(* IEC 61131-3 sources: plc-st-coding-agent/progress/evidence/f14_v11_public_20261113/jobs/custom_deepseek-v4pro (part 4) *)

(* ---- public-medium-02.raw_candidate_01.st ---- *)
TYPE ST_AnalogChannel :
STRUCT
    enable : BOOL;
    hiLIM : REAL;
    loLIM : REAL;
    bipolar : BOOL;
    measuringMode : INT;
    retVal : WORD;
    outputValue : REAL;
END_STRUCT
END_TYPE

FUNCTION_BLOCK AnalogBatchProcessing
VAR_INPUT
    count : DINT;
END_VAR
VAR_INOUT
    analogValues : ARRAY[*] OF INT;
    channels : ARRAY[*] OF ST_AnalogChannel;
END_VAR
VAR
    tmp_i : DINT;
    tmp_process_count : DINT;
    tmp_analog_lower : DINT;
    tmp_channel_lower : DINT;
    tmp_analog_len : DINT;
    tmp_channel_len : DINT;
    tmp_raw : INT;
    tmp_raw_real : REAL;
    tmp_span : REAL;
    tmp_range : REAL;
END_VAR

(* ENGINEERING_CONTRACT
   Outputs:
   channels[].retVal : activation = enabled channel processed; retention = written only then; reset = none; priority = mode error before limit error; units: WORD.
   channels[].outputValue : activation = successful conversion only; retention = unchanged on skip/error/disabled; reset = none; units: REAL.
   Disabled channels: no writes.
   Mode 0 scaling boundaries: unipolar raw 0..27648 maps [loLIM,hiLIM], bipolar raw -27648..27648 maps [loLIM,hiLIM]; no clamping specified (PUB003).
   Mode 1/2 scale raw/10, raw/100 (PUB004, PUB005).
   Count represents ordinal positions from each array lower bound; caller valid 0..min lengths (PUB001). Cap invalid high count to available.
   Priority for invalid mode vs limit: invalid mode 16#8001 checked first, then limit 16#8002 (PUB006, PUB007).
*)

(* CONTRACT_RULES [] *)

tmp_analog_lower := LOWER_BOUND(analogValues, 1);
tmp_channel_lower := LOWER_BOUND(channels, 1);
tmp_analog_len := UPPER_BOUND(analogValues, 1) - tmp_analog_lower + 1;
tmp_channel_len := UPPER_BOUND(channels, 1) - tmp_channel_lower + 1;

IF count <= 0 THEN
    RETURN;
END_IF;

tmp_process_count := count;
IF tmp_process_count > tmp_analog_len THEN
    tmp_process_count := tmp_analog_len;
END_IF;
IF tmp_process_count > tmp_channel_len THEN
    tmp_process_count := tmp_channel_len;
END_IF;

FOR tmp_i := 0 TO tmp_process_count - 1 DO
    IF channels[tmp_channel_lower + tmp_i].enable THEN
        IF channels[tmp_channel_lower + tmp_i].measuringMode < 0 OR
           channels[tmp_channel_lower + tmp_i].measuringMode > 2 THEN
            channels[tmp_channel_lower + tmp_i].retVal := 16#8001;
        ELSIF channels[tmp_channel_lower + tmp_i].hiLIM <= channels[tmp_channel_lower + tmp_i].loLIM THEN
            channels[tmp_channel_lower + tmp_i].retVal := 16#8002;
        ELSE
            channels[tmp_channel_lower + tmp_i].retVal := 0;
            tmp_raw := analogValues[tmp_analog_lower + tmp_i];
            tmp_raw_real := TO_REAL(tmp_raw);
            CASE channels[tmp_channel_lower + tmp_i].measuringMode OF
                0:
                    tmp_span := channels[tmp_channel_lower + tmp_i].hiLIM - channels[tmp_channel_lower + tmp_i].loLIM;
                    IF channels[tmp_channel_lower + tmp_i].bipolar THEN
                        tmp_range := 55296.0;
                        channels[tmp_channel_lower + tmp_i].outputValue :=
                            channels[tmp_channel_lower + tmp_i].loLIM +
                            ((tmp_raw_real + 27648.0) / tmp_range) * tmp_span;
                    ELSE
                        tmp_range := 27648.0;
                        channels[tmp_channel_lower + tmp_i].outputValue :=
                            channels[tmp_channel_lower + tmp_i].loLIM +
                            (tmp_raw_real / tmp_range) * tmp_span;
                    END_IF
                1:
                    channels[tmp_channel_lower + tmp_i].outputValue := tmp_raw_real / 10.0;
                2:
                    channels[tmp_channel_lower + tmp_i].outputValue := tmp_raw_real / 100.0;
            END_CASE
        END_IF
    END_IF
END_FOR

END_FUNCTION_BLOCK

(* ---- public-medium-02.raw_candidate_02.st ---- *)
TYPE ST_AnalogChannel :
STRUCT
    enable : BOOL;
    hiLIM : REAL;
    loLIM : REAL;
    bipolar : BOOL;
    measuringMode : INT;
    retVal : WORD;
    outputValue : REAL;
END_STRUCT
END_TYPE;

FUNCTION_BLOCK AnalogBatchProcessing
VAR_INPUT
    count : DINT;
END_VAR
VAR_IN_OUT
    analogValues : ARRAY[*] OF INT;
    channels : ARRAY[*] OF ST_AnalogChannel;
END_VAR
VAR
    tmp_i : DINT;
    tmp_process_count : DINT;
    tmp_analog_lower : DINT;
    tmp_channel_lower : DINT;
    tmp_analog_len : DINT;
    tmp_channel_len : DINT;
    tmp_raw : INT;
    tmp_raw_real : REAL;
    tmp_span : REAL;
    tmp_range : REAL;
END_VAR

(* ENGINEERING_CONTRACT
   Outputs:
   channels[].retVal : activation = enabled channel processed; retention = written only then; reset = none; priority = mode error before limit error; units: WORD.
   channels[].outputValue : activation = successful conversion only; retention = unchanged on skip/error/disabled; reset = none; units: REAL.
   Disabled channels: no writes.
   Mode 0 scaling boundaries: unipolar raw 0..27648 maps [loLIM,hiLIM], bipolar raw -27648..27648 maps [loLIM,hiLIM]; no clamping specified (PUB003).
   Mode 1/2 scale raw/10, raw/100 (PUB004, PUB005).
   Count represents ordinal positions from each array lower bound; caller valid 0..min lengths (PUB001). Cap invalid high count to available.
   Priority for invalid mode vs limit: invalid mode 16#8001 checked first, then limit 16#8002 (PUB006, PUB007).
*)

(* CONTRACT_RULES [] *)

tmp_analog_lower := LOWER_BOUND(analogValues, 1);
tmp_channel_lower := LOWER_BOUND(channels, 1);
tmp_analog_len := UPPER_BOUND(analogValues, 1) - tmp_analog_lower + 1;
tmp_channel_len := UPPER_BOUND(channels, 1) - tmp_channel_lower + 1;

IF count <= 0 THEN
    RETURN;
END_IF;

tmp_process_count := count;
IF tmp_process_count > tmp_analog_len THEN
    tmp_process_count := tmp_analog_len;
END_IF;
IF tmp_process_count > tmp_channel_len THEN
    tmp_process_count := tmp_channel_len;
END_IF;

FOR tmp_i := 0 TO tmp_process_count - 1 DO
    IF channels[tmp_channel_lower + tmp_i].enable THEN
        IF channels[tmp_channel_lower + tmp_i].measuringMode < 0 OR
           channels[tmp_channel_lower + tmp_i].measuringMode > 2 THEN
            channels[tmp_channel_lower + tmp_i].retVal := 16#8001;
        ELSIF channels[tmp_channel_lower + tmp_i].hiLIM <= channels[tmp_channel_lower + tmp_i].loLIM THEN
            channels[tmp_channel_lower + tmp_i].retVal := 16#8002;
        ELSE
            channels[tmp_channel_lower + tmp_i].retVal := 0;
            tmp_raw := analogValues[tmp_analog_lower + tmp_i];
            tmp_raw_real := TO_REAL(tmp_raw);
            CASE channels[tmp_channel_lower + tmp_i].measuringMode OF
                0:
                    tmp_span := channels[tmp_channel_lower + tmp_i].hiLIM - channels[tmp_channel_lower + tmp_i].loLIM;
                    IF channels[tmp_channel_lower + tmp_i].bipolar THEN
                        tmp_range := 55296.0;
                        channels[tmp_channel_lower + tmp_i].outputValue :=
                            channels[tmp_channel_lower + tmp_i].loLIM +
                            ((tmp_raw_real + 27648.0) / tmp_range) * tmp_span;
                    ELSE
                        tmp_range := 27648.0;
                        channels[tmp_channel_lower + tmp_i].outputValue :=
                            channels[tmp_channel_lower + tmp_i].loLIM +
                            (tmp_raw_real / tmp_range) * tmp_span;
                    END_IF;
                1:
                    channels[tmp_channel_lower + tmp_i].outputValue := tmp_raw_real / 10.0;
                2:
                    channels[tmp_channel_lower + tmp_i].outputValue := tmp_raw_real / 100.0;
            END_CASE;
        END_IF;
    END_IF;
END_FOR;

END_FUNCTION_BLOCK

(* ---- public-medium-03.candidate_01.st ---- *)
FUNCTION_BLOCK FB
VAR_INPUT
    cyclicExecution : BOOL;
    trigger : BOOL;
    value : LREAL;
    windowSize : INT;
    reset : BOOL;
END_VAR
VAR_OUTPUT
    average : LREAL;
    windowSizeReached : BOOL;
    error : BOOL;
    status : WORD;
END_VAR
VAR
    trig_rt : R_TRIG;
    buf : ARRAY[0..99] OF LREAL;
    head : INT := 0;
    count : INT := 0;
    n : INT;
    i : INT;
    idx : INT;
    do_update : BOOL;
    tmp_sum : LREAL;
    tmp_window_valid : BOOL;
END_VAR

(* ENGINEERING_CONTRACT
   - average: LREAL, updated only on new value read (cyclic scan or trigger rising edge while cyclicExecution FALSE);
     reset clears to 0.0. Unit: input value unit.
   - windowSizeReached: BOOL, TRUE iff count >= windowSize and window valid; reset clears; invalid window sets FALSE.
   - error/status: combinational; invalid window (windowSize < 1 or > 100) sets error TRUE, status 16#8200;
     otherwise error FALSE, status 16#0000.
   - reset has priority over read; invalid window blocks read and overrides status; no latch.
   - trigger rising edges are ignored while cyclicExecution TRUE.
   - circular buffer capacity 100; changing windowSize does not clear buffer.
*)
(* CONTRACT_RULES [] *)

trig_rt(CLK := trigger);
tmp_window_valid := (windowSize >= 1) AND (windowSize <= 100);

IF reset THEN
    head := 0;
    count := 0;
    average := 0.0;
    windowSizeReached := FALSE;

    IF tmp_window_valid THEN
        error := FALSE;
        status := WORD#16#0000;
    ELSE
        error := TRUE;
        status := WORD#16#8200;
    END_IF;
    RETURN;

ELSIF NOT tmp_window_valid THEN
    error := TRUE;
    status := WORD#16#8200;
    average := 0.0;
    windowSizeReached := FALSE;
    RETURN;

ELSE
    error := FALSE;
    status := WORD#16#0000;
    windowSizeReached := (count >= windowSize);

    do_update := FALSE;
    IF cyclicExecution THEN
        do_update := TRUE;
    ELSIF trig_rt.Q THEN
        do_update := TRUE;
    END_IF;

    IF do_update THEN
        buf[head] := value;
        head := (head + 1) MOD 100;
        IF count < 100 THEN
            count := count + 1;
        END_IF;

        n := count;
        IF n > windowSize THEN
            n := windowSize;
        END_IF;

        IF n = 0 THEN
            average := 0.0;
        ELSE
            tmp_sum := 0.0;
            FOR i := 0 TO n - 1 DO
                idx := (head - n + i) MOD 100;
                IF idx < 0 THEN
                    idx := idx + 100;
                END_IF;
                tmp_sum := tmp_sum + buf[idx];
            END_FOR;
            average := tmp_sum / INT_TO_LREAL(n);
        END_IF;

        windowSizeReached := (count >= windowSize);
    END_IF;
END_IF;

END_FUNCTION_BLOCK

(* ---- public-medium-03.raw_candidate_01.st ---- *)
FUNCTION_BLOCK FB
VAR_INPUT
    cyclicExecution : BOOL;
    trigger : BOOL;
    value : LREAL;
    windowSize : INT;
    reset : BOOL;
END_VAR
VAR_OUTPUT
    average : LREAL;
    windowSizeReached : BOOL;
    error : BOOL;
    status : WORD;
END_VAR
VAR
    trig_rt : R_TRIG;
    buf : ARRAY[0..99] OF LREAL;
    head : INT := 0;
    count : INT := 0;
    n : INT;
    i : INT;
    idx : INT;
    do_update : BOOL;
    tmp_sum : LREAL;
    tmp_window_valid : BOOL;
END_VAR

(* ENGINEERING_CONTRACT
   - average: LREAL, updated only on new value read (cyclic scan or trigger rising edge while cyclicExecution FALSE);
     reset clears to 0.0. Unit: input value unit.
   - windowSizeReached: BOOL, TRUE iff count >= windowSize and window valid; reset clears; invalid window sets FALSE.
   - error/status: combinational; invalid window (windowSize < 1 or > 100) sets error TRUE, status 16#8200;
     otherwise error FALSE, status 16#0000.
   - reset has priority over read; invalid window blocks read and overrides status; no latch.
   - trigger rising edges are ignored while cyclicExecution TRUE.
   - circular buffer capacity 100; changing windowSize does not clear buffer.
*)
(* CONTRACT_RULES [] *)

trig_rt(CLK := trigger);
tmp_window_valid := (windowSize >= 1) AND (windowSize <= 100);

IF reset THEN
    head := 0;
    count := 0;
    average := 0.0;
    windowSizeReached := FALSE;

    IF tmp_window_valid THEN
        error := FALSE;
        status := WORD#16#0000;
    ELSE
        error := TRUE;
        status := WORD#16#8200;
    END_IF;
    RETURN;

ELSIF NOT tmp_window_valid THEN
    error := TRUE;
    status := WORD#16#8200;
    average := 0.0;
    windowSizeReached := FALSE;
    RETURN;

ELSE
    error := FALSE;
    status := WORD#16#0000;
    windowSizeReached := (count >= windowSize);

    do_update := FALSE;
    IF cyclicExecution THEN
        do_update := TRUE;
    ELSIF trig_rt.Q THEN
        do_update := TRUE;
    END_IF;

    IF do_update THEN
        buf[head] := value;
        head := (head + 1) MOD 100;
        IF count < 100 THEN
            count := count + 1;
        END_IF;

        n := count;
        IF n > windowSize THEN
            n := windowSize;
        END_IF;

        IF n = 0 THEN
            average := 0.0;
        ELSE
            tmp_sum := 0.0;
            FOR i := 0 TO n - 1 DO
                idx := (head - n + i) MOD 100;
                IF idx < 0 THEN
                    idx := idx + 100;
                END_IF;
                tmp_sum := tmp_sum + buf[idx];
            END_FOR;
            average := tmp_sum / INT_TO_LREAL(n);
        END_IF;

        windowSizeReached := (count >= windowSize);
    END_IF;
END_IF;

END_FUNCTION_BLOCK

(* ---- public-medium-04.candidate_01.st ---- *)
FUNCTION_BLOCK FB_TemperatureControl
VAR_INPUT
    TemperatureSensorInput : REAL;
    SetTemperature : REAL;
END_VAR
VAR_OUTPUT
    CurrentTemperature : REAL;
    SetTempDisplay : REAL;
    HeaterStatus : BOOL;
    OverheatProtection : BOOL;
    HeaterOutput : BOOL;
END_VAR
VAR
    tmp_sensor_fault : BOOL;
    tmp_heat_allowed : BOOL;
    tmp_overheat_active : BOOL;
    tmp_heat_on_timer : TON;
    tmp_cooldown_timer : TON;
    tmp_heat_limit : TIME := T#5001MS;  (* strictly > 5 s continuous heating *)
    tmp_cooldown_limit : TIME := T#3S;
END_VAR

(*
ENGINEERING_CONTRACT
- CurrentTemperature/SetTempDisplay: combinational echoes, raw units.
- HeaterOutput: on when sensor valid, no overheat, sensor < set;
  off when sensor >= set, sensor fault, or overheat. Equal is off.
- OverheatProtection: latched TRUE on continuous heater on >5s; auto clear after 3s cooldown.
- HeaterStatus: echo of HeaterOutput.
- Sensor fault: <0.0 or >100.0. Fault and overheat force heater off.
- Unspecified: equal setpoint and reset after cooldown interpreted as above.
- PUB001-PUB008.
*)

(* CONTRACT_RULES [] *)

tmp_sensor_fault := (TemperatureSensorInput < 0.0) OR (TemperatureSensorInput > 100.0);

tmp_heat_allowed := (NOT tmp_sensor_fault)
                    AND (NOT tmp_overheat_active)
                    AND (TemperatureSensorInput < SetTemperature);

tmp_heat_on_timer(IN := tmp_heat_allowed, PT := tmp_heat_limit);

IF tmp_heat_on_timer.Q THEN
    tmp_overheat_active := TRUE;
END_IF;

tmp_cooldown_timer(IN := tmp_overheat_active, PT := tmp_cooldown_limit);

IF tmp_cooldown_timer.Q THEN
    tmp_overheat_active := FALSE;
END_IF;

HeaterOutput := (NOT tmp_sensor_fault)
                AND (NOT tmp_overheat_active)
                AND (TemperatureSensorInput < SetTemperature);

HeaterStatus := HeaterOutput;
OverheatProtection := tmp_overheat_active;
CurrentTemperature := TemperatureSensorInput;
SetTempDisplay := SetTemperature;

END_FUNCTION_BLOCK

(* ---- public-medium-04.candidate_02.st ---- *)
FUNCTION_BLOCK FB_TemperatureControl
VAR_INPUT
    TemperatureSensorInput : REAL;
    SetTemperature : REAL;
END_VAR
VAR_OUTPUT
    CurrentTemperature : REAL;
    SetTempDisplay : REAL;
    HeaterStatus : BOOL;
    OverheatProtection : BOOL;
    HeaterOutput : BOOL;
END_VAR
VAR
    tmp_sensor_fault : BOOL;
    tmp_heat_allowed : BOOL;
    tmp_overheat_active : BOOL;
    tmp_heat_on_timer : TON;
    tmp_cooldown_timer : TON;
    tmp_heat_limit : TIME := T#5001MS;  (* strictly > 5 s continuous heating *)
    tmp_cooldown_limit : TIME := T#3S;
END_VAR

(*
ENGINEERING_CONTRACT
- CurrentTemperature/SetTempDisplay: combinational echoes, raw units.
- HeaterOutput: on when sensor valid, no overheat, sensor < set;
  off when sensor >= set, sensor fault, or overheat. Equal is off.
- OverheatProtection: latched TRUE on continuous heater on >5s; auto clear after 3s cooldown.
- HeaterStatus: echo of HeaterOutput.
- Sensor fault: <0.0 or >100.0. Fault and overheat force heater off.
- Equal setpoint and reset after cooldown interpreted as above.
- Heat timer starts in same scan as heater is newly enabled; heat trip starts cooldown in same scan.
- PUB001-PUB008.
*)

(* CONTRACT_RULES [] *)

tmp_sensor_fault := (TemperatureSensorInput < 0.0) OR (TemperatureSensorInput > 100.0);

(* Process cooldown for any currently active overheat before computing heater command *)
tmp_cooldown_timer(IN := tmp_overheat_active, PT := tmp_cooldown_limit);
IF tmp_cooldown_timer.Q THEN
    tmp_overheat_active := FALSE;
END_IF;

tmp_heat_allowed := (NOT tmp_sensor_fault) AND (NOT tmp_overheat_active) AND (TemperatureSensorInput < SetTemperature);
HeaterOutput := tmp_heat_allowed;

tmp_heat_on_timer(IN := HeaterOutput, PT := tmp_heat_limit);
IF tmp_heat_on_timer.Q THEN
    tmp_overheat_active := TRUE;
    HeaterOutput := FALSE;
    (* Start cooldown timer on the same scan as the overheat trip *)
    tmp_cooldown_timer(IN := TRUE, PT := tmp_cooldown_limit);
END_IF;

HeaterStatus := HeaterOutput;
OverheatProtection := tmp_overheat_active;
CurrentTemperature := TemperatureSensorInput;
SetTempDisplay := SetTemperature;

END_FUNCTION_BLOCK

(* ---- public-medium-04.candidate_03.st ---- *)
FUNCTION_BLOCK FB_TemperatureControl
VAR_INPUT
    TemperatureSensorInput : REAL;
    SetTemperature : REAL;
END_VAR
VAR_OUTPUT
    CurrentTemperature : REAL;
    SetTempDisplay : REAL;
    HeaterStatus : BOOL;
    OverheatProtection : BOOL;
    HeaterOutput : BOOL;
END_VAR
VAR
    tmp_sensor_fault : BOOL;
    tmp_heat_allowed : BOOL;
    tmp_overheat_active : BOOL;
    tmp_heat_on_timer : TON;
    tmp_cooldown_timer : TON;
    tmp_heat_limit : TIME := T#5001MS;  (* strictly more than 5 s continuous heating *)
    tmp_cooldown_limit : TIME := T#3S;
END_VAR

(*
ENGINEERING_CONTRACT
- CurrentTemperature/SetTempDisplay are combinational echoes of the inputs.
- Sensor fault when input < 0.0 or > 100.0; fault forces heater off.
- HeaterOutput is on only when sensor valid, overheat protection inactive,
  and TemperatureSensorInput < SetTemperature. Equal setpoint is off.
- OverheatProtection latches when continuous heater-on time exceeds 5 s,
  and clears after a 3 s cooldown. Cooldown and same-scan reactivation are
  evaluated so clearing protection allows heater and its timer in the same scan.
- HeaterStatus follows HeaterOutput.
*)

(* CONTRACT_RULES [] *)

tmp_sensor_fault := (TemperatureSensorInput < 0.0) OR (TemperatureSensorInput > 100.0);

(* Evaluate cooldown first so a completed cooldown can lift protection
   and permit heater startup during this same invocation. *)
tmp_cooldown_timer(IN := tmp_overheat_active, PT := tmp_cooldown_limit);
IF tmp_cooldown_timer.Q THEN
    tmp_overheat_active := FALSE;
END_IF;

tmp_heat_allowed := (NOT tmp_sensor_fault)
                    AND (NOT tmp_overheat_active)
                    AND (TemperatureSensorInput < SetTemperature);

tmp_heat_on_timer(IN := tmp_heat_allowed, PT := tmp_heat_limit);

IF tmp_heat_on_timer.Q THEN
    tmp_overheat_active := TRUE;
    (* Start cooldown in the same scan when the overheat latch occurs. *)
    tmp_cooldown_timer(IN := TRUE, PT := tmp_cooldown_limit);
END_IF;

HeaterOutput := (NOT tmp_sensor_fault)
                AND (NOT tmp_overheat_active)
                AND (TemperatureSensorInput < SetTemperature);

HeaterStatus := HeaterOutput;
OverheatProtection := tmp_overheat_active;
CurrentTemperature := TemperatureSensorInput;
SetTempDisplay := SetTemperature;

END_FUNCTION_BLOCK

(* ---- public-medium-04.candidate_04.st ---- *)
FUNCTION_BLOCK FB_TemperatureControl
VAR_INPUT
    TemperatureSensorInput : REAL;
    SetTemperature : REAL;
END_VAR
VAR_OUTPUT
    CurrentTemperature : REAL;
    SetTempDisplay : REAL;
    HeaterStatus : BOOL;
    OverheatProtection : BOOL;
    HeaterOutput : BOOL;
END_VAR
VAR
    tmp_sensor_fault : BOOL;
    tmp_heat_allowed : BOOL;
    tmp_overheat_active : BOOL;
    tmp_heat_on_timer : TON;
    tmp_cooldown_timer : TON;
    tmp_heat_limit : TIME := T#5001MS;  (* strictly > 5 s continuous heating *)
    tmp_cooldown_limit : TIME := T#3S;
END_VAR

(*
ENGINEERING_CONTRACT
- CurrentTemperature/SetTempDisplay: combinational echoes, raw units.
- HeaterOutput: on when sensor valid, no overheat, sensor < set;
  off when sensor >= set, sensor fault, or overheat. Equal is off.
- OverheatProtection: latched TRUE on continuous heater on >5s; auto clear after 3s cooldown.
- HeaterStatus: echo of HeaterOutput.
- Sensor fault: <0.0 or >100.0. Fault and overheat force heater off.
- Unspecified: equal setpoint and reset after cooldown interpreted as above.
- PUB001-PUB008.
*)

(* CONTRACT_RULES [] *)

tmp_sensor_fault := (TemperatureSensorInput < 0.0) OR (TemperatureSensorInput > 100.0);

(* Cooldown logic first: if overheat is active and cooldown elapsed, clear it. *)
tmp_cooldown_timer(IN := tmp_overheat_active, PT := tmp_cooldown_limit);
IF tmp_cooldown_timer.Q THEN
    tmp_overheat_active := FALSE;
END_IF;

(* Recompute heater allowed using possibly updated overheat state. *)
tmp_heat_allowed := (NOT tmp_sensor_fault)
                    AND (NOT tmp_overheat_active)
                    AND (TemperatureSensorInput < SetTemperature);

(* Run heat timer after cooldown so it starts immediately when heater becomes allowed. *)
tmp_heat_on_timer(IN := tmp_heat_allowed, PT := tmp_heat_limit);
IF tmp_heat_on_timer.Q THEN
    tmp_overheat_active := TRUE;
END_IF;

HeaterOutput := (NOT tmp_sensor_fault)
                AND (NOT tmp_overheat_active)
                AND (TemperatureSensorInput < SetTemperature);

HeaterStatus := HeaterOutput;
OverheatProtection := tmp_overheat_active;
CurrentTemperature := TemperatureSensorInput;
SetTempDisplay := SetTemperature;

END_FUNCTION_BLOCK

(* ---- public-medium-04.raw_candidate_01.st ---- *)
FUNCTION_BLOCK FB_TemperatureControl
VAR_INPUT
    TemperatureSensorInput : REAL;
    SetTemperature : REAL;
END_VAR
VAR_OUTPUT
    CurrentTemperature : REAL;
    SetTempDisplay : REAL;
    HeaterStatus : BOOL;
    OverheatProtection : BOOL;
    HeaterOutput : BOOL;
END_VAR
VAR
    tmp_sensor_fault : BOOL;
    tmp_heat_allowed : BOOL;
    tmp_overheat_active : BOOL;
    tmp_heat_on_timer : TON;
    tmp_cooldown_timer : TON;
    tmp_heat_limit : TIME := T#5001MS;  (* strictly > 5 s continuous heating *)
    tmp_cooldown_limit : TIME := T#3S;
END_VAR

(*
ENGINEERING_CONTRACT
- CurrentTemperature/SetTempDisplay: combinational echoes, raw units.
- HeaterOutput: on when sensor valid, no overheat, sensor < set;
  off when sensor >= set, sensor fault, or overheat. Equal is off.
- OverheatProtection: latched TRUE on continuous heater on >5s; auto clear after 3s cooldown.
- HeaterStatus: echo of HeaterOutput.
- Sensor fault: <0.0 or >100.0. Fault and overheat force heater off.
- Unspecified: equal setpoint and reset after cooldown interpreted as above.
- PUB001-PUB008.
*)

(* CONTRACT_RULES [] *)

tmp_sensor_fault := (TemperatureSensorInput < 0.0) OR (TemperatureSensorInput > 100.0);

tmp_heat_allowed := (NOT tmp_sensor_fault)
                    AND (NOT tmp_overheat_active)
                    AND (TemperatureSensorInput < SetTemperature);

tmp_heat_on_timer(IN := tmp_heat_allowed, PT := tmp_heat_limit);

IF tmp_heat_on_timer.Q THEN
    tmp_overheat_active := TRUE;
END_IF;

tmp_cooldown_timer(IN := tmp_overheat_active, PT := tmp_cooldown_limit);

IF tmp_cooldown_timer.Q THEN
    tmp_overheat_active := FALSE;
END_IF;

HeaterOutput := (NOT tmp_sensor_fault)
                AND (NOT tmp_overheat_active)
                AND (TemperatureSensorInput < SetTemperature);

HeaterStatus := HeaterOutput;
OverheatProtection := tmp_overheat_active;
CurrentTemperature := TemperatureSensorInput;
SetTempDisplay := SetTemperature;

END_FUNCTION_BLOCK

(* ---- public-medium-04.raw_candidate_02.st ---- *)
FUNCTION_BLOCK FB_TemperatureControl
VAR_INPUT
    TemperatureSensorInput : REAL;
    SetTemperature : REAL;
END_VAR
VAR_OUTPUT
    CurrentTemperature : REAL;
    SetTempDisplay : REAL;
    HeaterStatus : BOOL;
    OverheatProtection : BOOL;
    HeaterOutput : BOOL;
END_VAR
VAR
    tmp_sensor_fault : BOOL;
    tmp_heat_allowed : BOOL;
    tmp_overheat_active : BOOL;
    tmp_heat_on_timer : TON;
    tmp_cooldown_timer : TON;
    tmp_heat_limit : TIME := T#5001MS;  (* strictly > 5 s continuous heating *)
    tmp_cooldown_limit : TIME := T#3S;
END_VAR

(*
ENGINEERING_CONTRACT
- CurrentTemperature/SetTempDisplay: combinational echoes, raw units.
- HeaterOutput: on when sensor valid, no overheat, sensor < set;
  off when sensor >= set, sensor fault, or overheat. Equal is off.
- OverheatProtection: latched TRUE on continuous heater on >5s; auto clear after 3s cooldown.
- HeaterStatus: echo of HeaterOutput.
- Sensor fault: <0.0 or >100.0. Fault and overheat force heater off.
- Equal setpoint and reset after cooldown interpreted as above.
- Heat timer starts in same scan as heater is newly enabled; heat trip starts cooldown in same scan.
- PUB001-PUB008.
*)

(* CONTRACT_RULES [] *)

tmp_sensor_fault := (TemperatureSensorInput < 0.0) OR (TemperatureSensorInput > 100.0);

(* Process cooldown for any currently active overheat before computing heater command *)
tmp_cooldown_timer(IN := tmp_overheat_active, PT := tmp_cooldown_limit);
IF tmp_cooldown_timer.Q THEN
    tmp_overheat_active := FALSE;
END_IF;

tmp_heat_allowed := (NOT tmp_sensor_fault) AND (NOT tmp_overheat_active) AND (TemperatureSensorInput < SetTemperature);
HeaterOutput := tmp_heat_allowed;

tmp_heat_on_timer(IN := HeaterOutput, PT := tmp_heat_limit);
IF tmp_heat_on_timer.Q THEN
    tmp_overheat_active := TRUE;
    HeaterOutput := FALSE;
    (* Start cooldown timer on the same scan as the overheat trip *)
    tmp_cooldown_timer(IN := TRUE, PT := tmp_cooldown_limit);
END_IF;

HeaterStatus := HeaterOutput;
OverheatProtection := tmp_overheat_active;
CurrentTemperature := TemperatureSensorInput;
SetTempDisplay := SetTemperature;

END_FUNCTION_BLOCK

(* ---- public-medium-04.raw_candidate_03.st ---- *)
FUNCTION_BLOCK FB_TemperatureControl
VAR_INPUT
    TemperatureSensorInput : REAL;
    SetTemperature : REAL;
END_VAR
VAR_OUTPUT
    CurrentTemperature : REAL;
    SetTempDisplay : REAL;
    HeaterStatus : BOOL;
    OverheatProtection : BOOL;
    HeaterOutput : BOOL;
END_VAR
VAR
    tmp_sensor_fault : BOOL;
    tmp_heat_allowed : BOOL;
    tmp_overheat_active : BOOL;
    tmp_heat_on_timer : TON;
    tmp_cooldown_timer : TON;
    tmp_heat_limit : TIME := T#5001MS;  (* strictly more than 5 s continuous heating *)
    tmp_cooldown_limit : TIME := T#3S;
END_VAR

(*
ENGINEERING_CONTRACT
- CurrentTemperature/SetTempDisplay are combinational echoes of the inputs.
- Sensor fault when input < 0.0 or > 100.0; fault forces heater off.
- HeaterOutput is on only when sensor valid, overheat protection inactive,
  and TemperatureSensorInput < SetTemperature. Equal setpoint is off.
- OverheatProtection latches when continuous heater-on time exceeds 5 s,
  and clears after a 3 s cooldown. Cooldown and same-scan reactivation are
  evaluated so clearing protection allows heater and its timer in the same scan.
- HeaterStatus follows HeaterOutput.
*)

(* CONTRACT_RULES [] *)

tmp_sensor_fault := (TemperatureSensorInput < 0.0) OR (TemperatureSensorInput > 100.0);

(* Evaluate cooldown first so a completed cooldown can lift protection
   and permit heater startup during this same invocation. *)
tmp_cooldown_timer(IN := tmp_overheat_active, PT := tmp_cooldown_limit);
IF tmp_cooldown_timer.Q THEN
    tmp_overheat_active := FALSE;
END_IF;

tmp_heat_allowed := (NOT tmp_sensor_fault)
                    AND (NOT tmp_overheat_active)
                    AND (TemperatureSensorInput < SetTemperature);

tmp_heat_on_timer(IN := tmp_heat_allowed, PT := tmp_heat_limit);

IF tmp_heat_on_timer.Q THEN
    tmp_overheat_active := TRUE;
    (* Start cooldown in the same scan when the overheat latch occurs. *)
    tmp_cooldown_timer(IN := TRUE, PT := tmp_cooldown_limit);
END_IF;

HeaterOutput := (NOT tmp_sensor_fault)
                AND (NOT tmp_overheat_active)
                AND (TemperatureSensorInput < SetTemperature);

HeaterStatus := HeaterOutput;
OverheatProtection := tmp_overheat_active;
CurrentTemperature := TemperatureSensorInput;
SetTempDisplay := SetTemperature;

END_FUNCTION_BLOCK

(* ---- public-medium-04.raw_candidate_04.st ---- *)
FUNCTION_BLOCK FB_TemperatureControl
VAR_INPUT
    TemperatureSensorInput : REAL;
    SetTemperature : REAL;
END_VAR
VAR_OUTPUT
    CurrentTemperature : REAL;
    SetTempDisplay : REAL;
    HeaterStatus : BOOL;
    OverheatProtection : BOOL;
    HeaterOutput : BOOL;
END_VAR
VAR
    tmp_sensor_fault : BOOL;
    tmp_heat_allowed : BOOL;
    tmp_overheat_active : BOOL;
    tmp_heat_on_timer : TON;
    tmp_cooldown_timer : TON;
    tmp_heat_limit : TIME := T#5001MS;  (* strictly > 5 s continuous heating *)
    tmp_cooldown_limit : TIME := T#3S;
END_VAR

(*
ENGINEERING_CONTRACT
- CurrentTemperature/SetTempDisplay: combinational echoes, raw units.
- HeaterOutput: on when sensor valid, no overheat, sensor < set;
  off when sensor >= set, sensor fault, or overheat. Equal is off.
- OverheatProtection: latched TRUE on continuous heater on >5s; auto clear after 3s cooldown.
- HeaterStatus: echo of HeaterOutput.
- Sensor fault: <0.0 or >100.0. Fault and overheat force heater off.
- Unspecified: equal setpoint and reset after cooldown interpreted as above.
- PUB001-PUB008.
*)

(* CONTRACT_RULES [] *)

tmp_sensor_fault := (TemperatureSensorInput < 0.0) OR (TemperatureSensorInput > 100.0);

(* Cooldown logic first: if overheat is active and cooldown elapsed, clear it. *)
tmp_cooldown_timer(IN := tmp_overheat_active, PT := tmp_cooldown_limit);
IF tmp_cooldown_timer.Q THEN
    tmp_overheat_active := FALSE;
END_IF;

(* Recompute heater allowed using possibly updated overheat state. *)
tmp_heat_allowed := (NOT tmp_sensor_fault)
                    AND (NOT tmp_overheat_active)
                    AND (TemperatureSensorInput < SetTemperature);

(* Run heat timer after cooldown so it starts immediately when heater becomes allowed. *)
tmp_heat_on_timer(IN := tmp_heat_allowed, PT := tmp_heat_limit);
IF tmp_heat_on_timer.Q THEN
    tmp_overheat_active := TRUE;
END_IF;

HeaterOutput := (NOT tmp_sensor_fault)
                AND (NOT tmp_overheat_active)
                AND (TemperatureSensorInput < SetTemperature);

HeaterStatus := HeaterOutput;
OverheatProtection := tmp_overheat_active;
CurrentTemperature := TemperatureSensorInput;
SetTempDisplay := SetTemperature;

END_FUNCTION_BLOCK

(* ---- public-medium-05.candidate_01.st ---- *)
(* ENGINEERING_CONTRACT
- Manual mode (Mode=FALSE): MotorForward set while ForwardButton AND NOT ReverseButton; MotorReverse set while ReverseButton AND NOT ForwardButton; simultaneous buttons deactivate both (PUB002).
- Automatic mode (Mode=TRUE): move_AB latch set by ButtonA R_TRIG while SensorA true; cleared when SensorB true. move_BC latch set by ButtonB R_TRIG while SensorB true; cleared when SensorC true.
- MotorForward = Mode AND (move_AB OR move_BC). MotorReverse is always FALSE in automatic mode (PUB003/PUB004).
- CompletionLight latch set by ButtonC R_TRIG while Mode=TRUE and SensorC true; held high; cleared when SensorC=FALSE regardless of Mode (PUB004).
- Same-scan priority: destination sensor clear wins over move set; simultaneous ForwardButton and ReverseButton -> both motor outputs FALSE.
*)

(* CONTRACT_RULES [] *)

FUNCTION_BLOCK ProductionLineControl
VAR_INPUT
    Mode : BOOL;
    ForwardButton : BOOL;
    ReverseButton : BOOL;
    SensorA : BOOL;
    SensorB : BOOL;
    SensorC : BOOL;
    ButtonA : BOOL;
    ButtonB : BOOL;
    ButtonC : BOOL;
END_VAR
VAR_OUTPUT
    MotorForward : BOOL;
    MotorReverse : BOOL;
    CompletionLight : BOOL;
END_VAR
VAR
    move_AB : BOOL := FALSE;
    move_BC : BOOL := FALSE;
    completion_latch : BOOL := FALSE;
    btnA_rt : R_TRIG;
    btnB_rt : R_TRIG;
    btnC_rt : R_TRIG;
END_VAR

btnA_rt(CLK := ButtonA);
btnB_rt(CLK := ButtonB);
btnC_rt(CLK := ButtonC);

IF Mode THEN
    IF btnA_rt.Q AND SensorA THEN
        move_AB := TRUE;
    END_IF;

    IF btnB_rt.Q AND SensorB THEN
        move_BC := TRUE;
    END_IF;

    IF btnC_rt.Q AND SensorC THEN
        completion_latch := TRUE;
    END_IF;
END_IF;

IF SensorB THEN
    move_AB := FALSE;
END_IF;

IF SensorC THEN
    move_BC := FALSE;
END_IF;

IF NOT SensorC THEN
    completion_latch := FALSE;
END_IF;

IF Mode THEN
    MotorForward := move_AB OR move_BC;
    MotorReverse := FALSE;
ELSE
    IF ForwardButton AND NOT ReverseButton THEN
        MotorForward := TRUE;
        MotorReverse := FALSE;
    ELSIF ReverseButton AND NOT ForwardButton THEN
        MotorForward := FALSE;
        MotorReverse := TRUE;
    ELSE
        MotorForward := FALSE;
        MotorReverse := FALSE;
    END_IF;
END_IF;

CompletionLight := completion_latch;

END_FUNCTION_BLOCK

(* ---- public-medium-05.candidate_02.st ---- *)
(* ENGINEERING_CONTRACT
- Manual mode (Mode=FALSE): MotorForward set while ForwardButton AND NOT ReverseButton; MotorReverse set while ReverseButton AND NOT ForwardButton; simultaneous buttons deactivate both (PUB002).
- Automatic mode (Mode=TRUE): move_AB latch set by ButtonA R_TRIG while SensorA true; cleared when SensorB true. move_BC latch set by ButtonB while SensorB true; cleared when SensorC true.
- MotorForward = Mode AND (move_AB OR move_BC). MotorReverse is always FALSE in automatic mode (PUB003/PUB004).
- CompletionLight latch set by ButtonC R_TRIG while Mode=TRUE and SensorC true; held high; cleared when SensorC=FALSE regardless of Mode (PUB004).
- Same-scan priority: destination sensor clear wins over move set; simultaneous ForwardButton and ReverseButton -> both motor outputs FALSE.
*)

(* CONTRACT_RULES [] *)

FUNCTION_BLOCK ProductionLineControl
VAR_INPUT
    Mode : BOOL;
    ForwardButton : BOOL;
    ReverseButton : BOOL;
    SensorA : BOOL;
    SensorB : BOOL;
    SensorC : BOOL;
    ButtonA : BOOL;
    ButtonB : BOOL;
    ButtonC : BOOL;
END_VAR
VAR_OUTPUT
    MotorForward : BOOL;
    MotorReverse : BOOL;
    CompletionLight : BOOL;
END_VAR
VAR
    move_AB : BOOL := FALSE;
    move_BC : BOOL := FALSE;
    completion_latch : BOOL := FALSE;
    btnA_rt : R_TRIG;
    btnB_rt : R_TRIG;
    btnC_rt : R_TRIG;
END_VAR

btnA_rt(CLK := ButtonA);
btnB_rt(CLK := ButtonB);
btnC_rt(CLK := ButtonC);

IF Mode THEN
    IF btnA_rt.Q AND SensorA THEN
        move_AB := TRUE;
    END_IF;

    IF ButtonB AND SensorB THEN
        move_BC := TRUE;
    END_IF;

    IF btnC_rt.Q AND SensorC THEN
        completion_latch := TRUE;
    END_IF;
END_IF;

IF SensorB THEN
    move_AB := FALSE;
END_IF;

IF SensorC THEN
    move_BC := FALSE;
END_IF;

IF NOT SensorC THEN
    completion_latch := FALSE;
END_IF;

IF Mode THEN
    MotorForward := move_AB OR move_BC;
    MotorReverse := FALSE;
ELSE
    IF ForwardButton AND NOT ReverseButton THEN
        MotorForward := TRUE;
        MotorReverse := FALSE;
    ELSIF ReverseButton AND NOT ForwardButton THEN
        MotorForward := FALSE;
        MotorReverse := TRUE;
    ELSE
        MotorForward := FALSE;
        MotorReverse := FALSE;
    END_IF;
END_IF;

CompletionLight := completion_latch;

END_FUNCTION_BLOCK

(* ---- public-medium-05.candidate_03.st ---- *)
(* ENGINEERING_CONTRACT
- Manual mode (Mode=FALSE): MotorForward set while ForwardButton AND NOT ReverseButton; MotorReverse set while ReverseButton AND NOT ForwardButton; simultaneous buttons deactivate both (PUB002).
- Automatic mode (Mode=TRUE): move_AB latch set by ButtonA R_TRIG while SensorA true; cleared when SensorB true. move_BC latch set by ButtonB while SensorB true; cleared when SensorC true.
- MotorForward = Mode AND (move_AB OR move_BC). MotorReverse is always FALSE in automatic mode (PUB003/PUB004).
- CompletionLight latch set by ButtonC R_TRIG while Mode=TRUE and SensorC true; held high; cleared when SensorC=FALSE regardless of Mode (PUB004).
- Same-scan priority: destination sensor clear wins over move set; simultaneous ForwardButton and ReverseButton -> both motor outputs FALSE.
*)

(* CONTRACT_RULES [] *)

FUNCTION_BLOCK ProductionLineControl
VAR_INPUT
    Mode : BOOL;
    ForwardButton : BOOL;
    ReverseButton : BOOL;
    SensorA : BOOL;
    SensorB : BOOL;
    SensorC : BOOL;
    ButtonA : BOOL;
    ButtonB : BOOL;
    ButtonC : BOOL;
END_VAR
VAR_OUTPUT
    MotorForward : BOOL;
    MotorReverse : BOOL;
    CompletionLight : BOOL;
END_VAR
VAR
    move_AB : BOOL := FALSE;
    move_BC : BOOL := FALSE;
    completion_latch : BOOL := FALSE;
    btnA_rt : R_TRIG;
    btnB_rt : R_TRIG;
    btnC_rt : R_TRIG;
END_VAR

btnA_rt(CLK := ButtonA);
btnB_rt(CLK := ButtonB);
btnC_rt(CLK := ButtonC);

IF Mode THEN
    IF btnA_rt.Q AND SensorA THEN
        move_AB := TRUE;
    END_IF;

    IF btnB_rt.Q AND SensorB THEN
        move_BC := TRUE;
    END_IF;

    IF btnC_rt.Q AND SensorC THEN
        completion_latch := TRUE;
    END_IF;
END_IF;

IF SensorB THEN
    move_AB := FALSE;
END_IF;

IF SensorC THEN
    move_BC := FALSE;
END_IF;

IF NOT SensorC THEN
    completion_latch := FALSE;
END_IF;

IF Mode THEN
    MotorForward := move_AB OR move_BC;
    MotorReverse := FALSE;
ELSE
    IF ForwardButton AND NOT ReverseButton THEN
        MotorForward := TRUE;
        MotorReverse := FALSE;
    ELSIF ReverseButton AND NOT ForwardButton THEN
        MotorForward := FALSE;
        MotorReverse := TRUE;
    ELSE
        MotorForward := FALSE;
        MotorReverse := FALSE;
    END_IF;
END_IF;

CompletionLight := completion_latch;

END_FUNCTION_BLOCK

(* ---- public-medium-05.candidate_04.st ---- *)
(* ENGINEERING_CONTRACT
- Manual mode (Mode=FALSE): MotorForward set while ForwardButton AND NOT ReverseButton; MotorReverse set while ReverseButton AND NOT ForwardButton; simultaneous buttons deactivate both (PUB002).
- Automatic mode (Mode=TRUE): move_AB latch set by ButtonA R_TRIG while SensorA true; cleared when SensorB true. move_BC latch set by ButtonB R_TRIG while SensorB true; cleared when SensorC true.
- MotorForward = Mode AND (move_AB OR move_BC). MotorReverse is always FALSE in automatic mode (PUB003/PUB004).
- CompletionLight latch set by ButtonC R_TRIG while Mode=TRUE and SensorC true; held high; cleared when SensorC=FALSE regardless of Mode (PUB004).
- Same-scan priority: destination sensor clear wins over move set; simultaneous ForwardButton and ReverseButton -> both motor outputs FALSE.
*)

(* CONTRACT_RULES [] *)

FUNCTION_BLOCK ProductionLineControl
VAR_INPUT
    Mode : BOOL;
    ForwardButton : BOOL;
    ReverseButton : BOOL;
    SensorA : BOOL;
    SensorB : BOOL;
    SensorC : BOOL;
    ButtonA : BOOL;
    ButtonB : BOOL;
    ButtonC : BOOL;
END_VAR
VAR_OUTPUT
    MotorForward : BOOL;
    MotorReverse : BOOL;
    CompletionLight : BOOL;
END_VAR
VAR
    move_AB : BOOL := FALSE;
    move_BC : BOOL := FALSE;
    completion_latch : BOOL := FALSE;
    btnA_rt : R_TRIG;
    btnB_rt : R_TRIG;
    btnC_rt : R_TRIG;
END_VAR

btnA_rt(CLK := ButtonA);
btnB_rt(CLK := ButtonB);
btnC_rt(CLK := ButtonC);

IF Mode THEN
    IF btnA_rt.Q AND SensorA THEN
        move_AB := TRUE;
    END_IF;

    IF btnB_rt.Q AND SensorB THEN
        move_BC := TRUE;
    END_IF;

    IF btnC_rt.Q AND SensorC THEN
        completion_latch := TRUE;
    END_IF;
END_IF;

IF SensorB THEN
    move_AB := FALSE;
END_IF;

IF SensorC THEN
    move_BC := FALSE;
END_IF;

IF NOT SensorC THEN
    completion_latch := FALSE;
END_IF;

IF Mode THEN
    MotorForward := move_AB OR move_BC;
    MotorReverse := FALSE;
ELSE
    IF ForwardButton AND NOT ReverseButton THEN
        MotorForward := TRUE;
        MotorReverse := FALSE;
    ELSIF ReverseButton AND NOT ForwardButton THEN
        MotorForward := FALSE;
        MotorReverse := TRUE;
    ELSE
        MotorForward := FALSE;
        MotorReverse := FALSE;
    END_IF;
END_IF;

CompletionLight := completion_latch;

END_FUNCTION_BLOCK

(* ---- public-medium-05.raw_candidate_01.st ---- *)
(* ENGINEERING_CONTRACT
- Manual mode (Mode=FALSE): MotorForward set while ForwardButton AND NOT ReverseButton; MotorReverse set while ReverseButton AND NOT ForwardButton; simultaneous buttons deactivate both (PUB002).
- Automatic mode (Mode=TRUE): move_AB latch set by ButtonA R_TRIG while SensorA true; cleared when SensorB true. move_BC latch set by ButtonB R_TRIG while SensorB true; cleared when SensorC true.
- MotorForward = Mode AND (move_AB OR move_BC). MotorReverse is always FALSE in automatic mode (PUB003/PUB004).
- CompletionLight latch set by ButtonC R_TRIG while Mode=TRUE and SensorC true; held high; cleared when SensorC=FALSE regardless of Mode (PUB004).
- Same-scan priority: destination sensor clear wins over move set; simultaneous ForwardButton and ReverseButton -> both motor outputs FALSE.
*)

(* CONTRACT_RULES [] *)

FUNCTION_BLOCK ProductionLineControl
VAR_INPUT
    Mode : BOOL;
    ForwardButton : BOOL;
    ReverseButton : BOOL;
    SensorA : BOOL;
    SensorB : BOOL;
    SensorC : BOOL;
    ButtonA : BOOL;
    ButtonB : BOOL;
    ButtonC : BOOL;
END_VAR
VAR_OUTPUT
    MotorForward : BOOL;
    MotorReverse : BOOL;
    CompletionLight : BOOL;
END_VAR
VAR
    move_AB : BOOL := FALSE;
    move_BC : BOOL := FALSE;
    completion_latch : BOOL := FALSE;
    btnA_rt : R_TRIG;
    btnB_rt : R_TRIG;
    btnC_rt : R_TRIG;
END_VAR

btnA_rt(CLK := ButtonA);
btnB_rt(CLK := ButtonB);
btnC_rt(CLK := ButtonC);

IF Mode THEN
    IF btnA_rt.Q AND SensorA THEN
        move_AB := TRUE;
    END_IF;

    IF btnB_rt.Q AND SensorB THEN
        move_BC := TRUE;
    END_IF;

    IF btnC_rt.Q AND SensorC THEN
        completion_latch := TRUE;
    END_IF;
END_IF;

IF SensorB THEN
    move_AB := FALSE;
END_IF;

IF SensorC THEN
    move_BC := FALSE;
END_IF;

IF NOT SensorC THEN
    completion_latch := FALSE;
END_IF;

IF Mode THEN
    MotorForward := move_AB OR move_BC;
    MotorReverse := FALSE;
ELSE
    IF ForwardButton AND NOT ReverseButton THEN
        MotorForward := TRUE;
        MotorReverse := FALSE;
    ELSIF ReverseButton AND NOT ForwardButton THEN
        MotorForward := FALSE;
        MotorReverse := TRUE;
    ELSE
        MotorForward := FALSE;
        MotorReverse := FALSE;
    END_IF;
END_IF;

CompletionLight := completion_latch;

END_FUNCTION_BLOCK

(* ---- public-medium-05.raw_candidate_02.st ---- *)
(* ENGINEERING_CONTRACT
- Manual mode (Mode=FALSE): MotorForward set while ForwardButton AND NOT ReverseButton; MotorReverse set while ReverseButton AND NOT ForwardButton; simultaneous buttons deactivate both (PUB002).
- Automatic mode (Mode=TRUE): move_AB latch set by ButtonA R_TRIG while SensorA true; cleared when SensorB true. move_BC latch set by ButtonB while SensorB true; cleared when SensorC true.
- MotorForward = Mode AND (move_AB OR move_BC). MotorReverse is always FALSE in automatic mode (PUB003/PUB004).
- CompletionLight latch set by ButtonC R_TRIG while Mode=TRUE and SensorC true; held high; cleared when SensorC=FALSE regardless of Mode (PUB004).
- Same-scan priority: destination sensor clear wins over move set; simultaneous ForwardButton and ReverseButton -> both motor outputs FALSE.
*)

(* CONTRACT_RULES [] *)

FUNCTION_BLOCK ProductionLineControl
VAR_INPUT
    Mode : BOOL;
    ForwardButton : BOOL;
    ReverseButton : BOOL;
    SensorA : BOOL;
    SensorB : BOOL;
    SensorC : BOOL;
    ButtonA : BOOL;
    ButtonB : BOOL;
    ButtonC : BOOL;
END_VAR
VAR_OUTPUT
    MotorForward : BOOL;
    MotorReverse : BOOL;
    CompletionLight : BOOL;
END_VAR
VAR
    move_AB : BOOL := FALSE;
    move_BC : BOOL := FALSE;
    completion_latch : BOOL := FALSE;
    btnA_rt : R_TRIG;
    btnB_rt : R_TRIG;
    btnC_rt : R_TRIG;
END_VAR

btnA_rt(CLK := ButtonA);
btnB_rt(CLK := ButtonB);
btnC_rt(CLK := ButtonC);

IF Mode THEN
    IF btnA_rt.Q AND SensorA THEN
        move_AB := TRUE;
    END_IF;

    IF ButtonB AND SensorB THEN
        move_BC := TRUE;
    END_IF;

    IF btnC_rt.Q AND SensorC THEN
        completion_latch := TRUE;
    END_IF;
END_IF;

IF SensorB THEN
    move_AB := FALSE;
END_IF;

IF SensorC THEN
    move_BC := FALSE;
END_IF;

IF NOT SensorC THEN
    completion_latch := FALSE;
END_IF;

IF Mode THEN
    MotorForward := move_AB OR move_BC;
    MotorReverse := FALSE;
ELSE
    IF ForwardButton AND NOT ReverseButton THEN
        MotorForward := TRUE;
        MotorReverse := FALSE;
    ELSIF ReverseButton AND NOT ForwardButton THEN
        MotorForward := FALSE;
        MotorReverse := TRUE;
    ELSE
        MotorForward := FALSE;
        MotorReverse := FALSE;
    END_IF;
END_IF;

CompletionLight := completion_latch;

END_FUNCTION_BLOCK

(* ---- public-medium-05.raw_candidate_03.st ---- *)
(* ENGINEERING_CONTRACT
- Manual mode (Mode=FALSE): MotorForward set while ForwardButton AND NOT ReverseButton; MotorReverse set while ReverseButton AND NOT ForwardButton; simultaneous buttons deactivate both (PUB002).
- Automatic mode (Mode=TRUE): move_AB latch set by ButtonA R_TRIG while SensorA true; cleared when SensorB true. move_BC latch set by ButtonB while SensorB true; cleared when SensorC true.
- MotorForward = Mode AND (move_AB OR move_BC). MotorReverse is always FALSE in automatic mode (PUB003/PUB004).
- CompletionLight latch set by ButtonC R_TRIG while Mode=TRUE and SensorC true; held high; cleared when SensorC=FALSE regardless of Mode (PUB004).
- Same-scan priority: destination sensor clear wins over move set; simultaneous ForwardButton and ReverseButton -> both motor outputs FALSE.
*)

(* CONTRACT_RULES [] *)

FUNCTION_BLOCK ProductionLineControl
VAR_INPUT
    Mode : BOOL;
    ForwardButton : BOOL;
    ReverseButton : BOOL;
    SensorA : BOOL;
    SensorB : BOOL;
    SensorC : BOOL;
    ButtonA : BOOL;
    ButtonB : BOOL;
    ButtonC : BOOL;
END_VAR
VAR_OUTPUT
    MotorForward : BOOL;
    MotorReverse : BOOL;
    CompletionLight : BOOL;
END_VAR
VAR
    move_AB : BOOL := FALSE;
    move_BC : BOOL := FALSE;
    completion_latch : BOOL := FALSE;
    btnA_rt : R_TRIG;
    btnB_rt : R_TRIG;
    btnC_rt : R_TRIG;
END_VAR

btnA_rt(CLK := ButtonA);
btnB_rt(CLK := ButtonB);
btnC_rt(CLK := ButtonC);

IF Mode THEN
    IF btnA_rt.Q AND SensorA THEN
        move_AB := TRUE;
    END_IF;

    IF btnB_rt.Q AND SensorB THEN
        move_BC := TRUE;
    END_IF;

    IF btnC_rt.Q AND SensorC THEN
        completion_latch := TRUE;
    END_IF;
END_IF;

IF SensorB THEN
    move_AB := FALSE;
END_IF;

IF SensorC THEN
    move_BC := FALSE;
END_IF;

IF NOT SensorC THEN
    completion_latch := FALSE;
END_IF;

IF Mode THEN
    MotorForward := move_AB OR move_BC;
    MotorReverse := FALSE;
ELSE
    IF ForwardButton AND NOT ReverseButton THEN
        MotorForward := TRUE;
        MotorReverse := FALSE;
    ELSIF ReverseButton AND NOT ForwardButton THEN
        MotorForward := FALSE;
        MotorReverse := TRUE;
    ELSE
        MotorForward := FALSE;
        MotorReverse := FALSE;
    END_IF;
END_IF;

CompletionLight := completion_latch;

END_FUNCTION_BLOCK

(* ---- public-medium-05.raw_candidate_04.st ---- *)
(* ENGINEERING_CONTRACT
- Manual mode (Mode=FALSE): MotorForward set while ForwardButton AND NOT ReverseButton; MotorReverse set while ReverseButton AND NOT ForwardButton; simultaneous buttons deactivate both (PUB002).
- Automatic mode (Mode=TRUE): move_AB latch set by ButtonA R_TRIG while SensorA true; cleared when SensorB true. move_BC latch set by ButtonB R_TRIG while SensorB true; cleared when SensorC true.
- MotorForward = Mode AND (move_AB OR move_BC). MotorReverse is always FALSE in automatic mode (PUB003/PUB004).
- CompletionLight latch set by ButtonC R_TRIG while Mode=TRUE and SensorC true; held high; cleared when SensorC=FALSE regardless of Mode (PUB004).
- Same-scan priority: destination sensor clear wins over move set; simultaneous ForwardButton and ReverseButton -> both motor outputs FALSE.
*)

(* CONTRACT_RULES [] *)

FUNCTION_BLOCK ProductionLineControl
VAR_INPUT
    Mode : BOOL;
    ForwardButton : BOOL;
    ReverseButton : BOOL;
    SensorA : BOOL;
    SensorB : BOOL;
    SensorC : BOOL;
    ButtonA : BOOL;
    ButtonB : BOOL;
    ButtonC : BOOL;
END_VAR
VAR_OUTPUT
    MotorForward : BOOL;
    MotorReverse : BOOL;
    CompletionLight : BOOL;
END_VAR
VAR
    move_AB : BOOL := FALSE;
    move_BC : BOOL := FALSE;
    completion_latch : BOOL := FALSE;
    btnA_rt : R_TRIG;
    btnB_rt : R_TRIG;
    btnC_rt : R_TRIG;
END_VAR

btnA_rt(CLK := ButtonA);
btnB_rt(CLK := ButtonB);
btnC_rt(CLK := ButtonC);

IF Mode THEN
    IF btnA_rt.Q AND SensorA THEN
        move_AB := TRUE;
    END_IF;

    IF btnB_rt.Q AND SensorB THEN
        move_BC := TRUE;
    END_IF;

    IF btnC_rt.Q AND SensorC THEN
        completion_latch := TRUE;
    END_IF;
END_IF;

IF SensorB THEN
    move_AB := FALSE;
END_IF;

IF SensorC THEN
    move_BC := FALSE;
END_IF;

IF NOT SensorC THEN
    completion_latch := FALSE;
END_IF;

IF Mode THEN
    MotorForward := move_AB OR move_BC;
    MotorReverse := FALSE;
ELSE
    IF ForwardButton AND NOT ReverseButton THEN
        MotorForward := TRUE;
        MotorReverse := FALSE;
    ELSIF ReverseButton AND NOT ForwardButton THEN
        MotorForward := FALSE;
        MotorReverse := TRUE;
    ELSE
        MotorForward := FALSE;
        MotorReverse := FALSE;
    END_IF;
END_IF;

CompletionLight := completion_latch;

END_FUNCTION_BLOCK

(* ---- public-medium-06.candidate_01.st ---- *)
FUNCTION_BLOCK SlabThicknessAlarmFaultHistory
VAR_INPUT
    THICKNESS_FAULT : BOOL;
    THICKNESS_SIGNAL_VALID : BOOL;
    CUTTING_RUN : BOOL;
    FaultTimestamp : DINT;
    CycleTime : TIME;
END_VAR
VAR_OUTPUT
    THICKNESS_ALARM : BOOL;
    Slab_Fault_Counter : UINT;
    Slab_Runtime_Accumulator : LTIME;
    Slab_Fault_History : ARRAY[0..4] OF DINT;
END_VAR
VAR
    alarm_hold : BOOL := FALSE;
    alarm_timer : TON;
    prev_valid_fault : BOOL := FALSE;
    init_done : BOOL := FALSE;
    valid_fault : BOOL;
END_VAR

(* ENGINEERING_CONTRACT
   THICKNESS_ALARM: set when valid_fault TRUE; hold after fault deassert until 500ms TON.Q;
   clear on signal invalid or power-up; invalid signal has same-scan priority; PUB001/PUB004.
   Slab_Fault_Counter: increments on valid_fault FALSE->TRUE; power-up zero; UINT count; PUB002/PUB005.
   Slab_Runtime_Accumulator: adds CycleTime only while valid, CUTTING_RUN and no fault;
   preserved otherwise; power-up zero; LTIME ns; PUB003/PUB004/PUB005.
   Slab_Fault_History: index 0 newest; shifted right on fault edge; power-up all zero;
   DINT seconds per FaultTimestamp; PUB002/PUB005/PUB006.
   Alarm hold timer restarts on each fault deassert while signal remains valid; PUB001.
   Unspecified: UINT rollover behavior interpreted as natural wrap; PUB006.
*)
(* CONTRACT_RULES [] *)

valid_fault := THICKNESS_SIGNAL_VALID AND THICKNESS_FAULT;

IF NOT init_done THEN
    init_done := TRUE;
    prev_valid_fault := valid_fault;
    Slab_Fault_Counter := UINT#0;
    Slab_Runtime_Accumulator := LTIME#0s;
    Slab_Fault_History[0] := DINT#0;
    Slab_Fault_History[1] := DINT#0;
    Slab_Fault_History[2] := DINT#0;
    Slab_Fault_History[3] := DINT#0;
    Slab_Fault_History[4] := DINT#0;
    alarm_hold := FALSE;
    alarm_timer(IN := FALSE, PT := T#500MS);
    THICKNESS_ALARM := FALSE;
ELSE
    IF valid_fault AND NOT prev_valid_fault THEN
        Slab_Fault_History[4] := Slab_Fault_History[3];
        Slab_Fault_History[3] := Slab_Fault_History[2];
        Slab_Fault_History[2] := Slab_Fault_History[1];
        Slab_Fault_History[1] := Slab_Fault_History[0];
        Slab_Fault_History[0] := FaultTimestamp;
        Slab_Fault_Counter := Slab_Fault_Counter + UINT#1;
    END_IF;

    prev_valid_fault := valid_fault;

    IF valid_fault THEN
        alarm_hold := TRUE;
    ELSIF NOT THICKNESS_SIGNAL_VALID THEN
        alarm_hold := FALSE;
    ELSIF alarm_timer.Q THEN
        alarm_hold := FALSE;
    END_IF;

    alarm_timer(IN := THICKNESS_SIGNAL_VALID AND NOT THICKNESS_FAULT, PT := T#500MS);

    THICKNESS_ALARM := THICKNESS_SIGNAL_VALID AND (valid_fault OR alarm_hold);

    IF THICKNESS_SIGNAL_VALID AND CUTTING_RUN AND NOT THICKNESS_FAULT AND (CycleTime > T#0ms) THEN
        Slab_Runtime_Accumulator := Slab_Runtime_Accumulator + TO_LTIME(CycleTime);
    END_IF;
END_IF;
END_FUNCTION_BLOCK

(* ---- public-medium-06.candidate_02.st ---- *)
(* ENGINEERING_CONTRACT
   THICKNESS_ALARM: latch on valid-fault FALSE->TRUE edge; hold via alarm_hold until TON reaches PT after fault deassert;
   clear on signal invalid; output = signal valid AND alarm_hold; PUB001/PUB004. Current TON.Q read after call.
   Slab_Fault_Counter: increment on same edge; wrap at UINT natural boundary; PUB002/PUB005.
   Slab_Runtime_Accumulator: add TO_LTIME(CycleTime) when valid and CUTTING_RUN and no fault and CycleTime>0 including first scan; LTIME ns; PUB003/PUB004.
   Slab_Fault_History[0..4]: shift oldest right, store timestamp at index0; PUB002/PUB006.
   Power-up: clear all stored state then process current inputs; prev_valid_fault starts false so first valid fault is a transition; PUB005.
   Unspecified: initial fault + invalid signal keeps alarm off until next edge; PUB004/PUB006.
*)
(* CONTRACT_RULES [] *)
FUNCTION_BLOCK SlabThicknessAlarmFaultHistory
VAR_INPUT
    THICKNESS_FAULT : BOOL;
    THICKNESS_SIGNAL_VALID : BOOL;
    CUTTING_RUN : BOOL;
    FaultTimestamp : DINT;
    CycleTime : TIME;
END_VAR
VAR_OUTPUT
    THICKNESS_ALARM : BOOL;
    Slab_Fault_Counter : UINT;
    Slab_Runtime_Accumulator : LTIME;
    Slab_Fault_History : ARRAY[0..4] OF DINT;
END_VAR
VAR
    alarm_hold : BOOL := FALSE;
    alarm_timer : TON;
    prev_valid_fault : BOOL := FALSE;
    init_done : BOOL := FALSE;
    valid_fault : BOOL;
END_VAR

valid_fault := THICKNESS_SIGNAL_VALID AND THICKNESS_FAULT;

IF NOT init_done THEN
    init_done := TRUE;
    Slab_Fault_Counter := UINT#0;
    Slab_Runtime_Accumulator := LTIME#0s;
    Slab_Fault_History[0] := DINT#0;
    Slab_Fault_History[1] := DINT#0;
    Slab_Fault_History[2] := DINT#0;
    Slab_Fault_History[3] := DINT#0;
    Slab_Fault_History[4] := DINT#0;
    alarm_hold := FALSE;
    alarm_timer(IN := FALSE, PT := T#500MS);
    THICKNESS_ALARM := FALSE;
END_IF;

IF valid_fault AND NOT prev_valid_fault THEN
    Slab_Fault_History[4] := Slab_Fault_History[3];
    Slab_Fault_History[3] := Slab_Fault_History[2];
    Slab_Fault_History[2] := Slab_Fault_History[1];
    Slab_Fault_History[1] := Slab_Fault_History[0];
    Slab_Fault_History[0] := FaultTimestamp;
    Slab_Fault_Counter := Slab_Fault_Counter + UINT#1;
    alarm_hold := TRUE;
END_IF;

prev_valid_fault := valid_fault;

alarm_timer(IN := THICKNESS_SIGNAL_VALID AND NOT THICKNESS_FAULT, PT := T#500MS);

IF NOT THICKNESS_SIGNAL_VALID THEN
    alarm_hold := FALSE;
ELSIF NOT valid_fault AND alarm_timer.Q THEN
    alarm_hold := FALSE;
END_IF;

THICKNESS_ALARM := THICKNESS_SIGNAL_VALID AND alarm_hold;

IF THICKNESS_SIGNAL_VALID AND CUTTING_RUN AND NOT THICKNESS_FAULT AND (CycleTime > T#0ms) THEN
    Slab_Runtime_Accumulator := Slab_Runtime_Accumulator + TO_LTIME(CycleTime);
END_IF;

END_FUNCTION_BLOCK

(* ---- public-medium-06.raw_candidate_01.st ---- *)
FUNCTION_BLOCK SlabThicknessAlarmFaultHistory
VAR_INPUT
    THICKNESS_FAULT : BOOL;
    THICKNESS_SIGNAL_VALID : BOOL;
    CUTTING_RUN : BOOL;
    FaultTimestamp : DINT;
    CycleTime : TIME;
END_VAR
VAR_OUTPUT
    THICKNESS_ALARM : BOOL;
    Slab_Fault_Counter : UINT;
    Slab_Runtime_Accumulator : LTIME;
    Slab_Fault_History : ARRAY[0..4] OF DINT;
END_VAR
VAR
    alarm_hold : BOOL := FALSE;
    alarm_timer : TON;
    prev_valid_fault : BOOL := FALSE;
    init_done : BOOL := FALSE;
    valid_fault : BOOL;
END_VAR

(* ENGINEERING_CONTRACT
   THICKNESS_ALARM: set when valid_fault TRUE; hold after fault deassert until 500ms TON.Q;
   clear on signal invalid or power-up; invalid signal has same-scan priority; PUB001/PUB004.
   Slab_Fault_Counter: increments on valid_fault FALSE->TRUE; power-up zero; UINT count; PUB002/PUB005.
   Slab_Runtime_Accumulator: adds CycleTime only while valid, CUTTING_RUN and no fault;
   preserved otherwise; power-up zero; LTIME ns; PUB003/PUB004/PUB005.
   Slab_Fault_History: index 0 newest; shifted right on fault edge; power-up all zero;
   DINT seconds per FaultTimestamp; PUB002/PUB005/PUB006.
   Alarm hold timer restarts on each fault deassert while signal remains valid; PUB001.
   Unspecified: UINT rollover behavior interpreted as natural wrap; PUB006.
*)
(* CONTRACT_RULES [] *)

valid_fault := THICKNESS_SIGNAL_VALID AND THICKNESS_FAULT;

IF NOT init_done THEN
    init_done := TRUE;
    prev_valid_fault := valid_fault;
    Slab_Fault_Counter := UINT#0;
    Slab_Runtime_Accumulator := LTIME#0s;
    Slab_Fault_History[0] := DINT#0;
    Slab_Fault_History[1] := DINT#0;
    Slab_Fault_History[2] := DINT#0;
    Slab_Fault_History[3] := DINT#0;
    Slab_Fault_History[4] := DINT#0;
    alarm_hold := FALSE;
    alarm_timer(IN := FALSE, PT := T#500MS);
    THICKNESS_ALARM := FALSE;
ELSE
    IF valid_fault AND NOT prev_valid_fault THEN
        Slab_Fault_History[4] := Slab_Fault_History[3];
        Slab_Fault_History[3] := Slab_Fault_History[2];
        Slab_Fault_History[2] := Slab_Fault_History[1];
        Slab_Fault_History[1] := Slab_Fault_History[0];
        Slab_Fault_History[0] := FaultTimestamp;
        Slab_Fault_Counter := Slab_Fault_Counter + UINT#1;
    END_IF;

    prev_valid_fault := valid_fault;

    IF valid_fault THEN
        alarm_hold := TRUE;
    ELSIF NOT THICKNESS_SIGNAL_VALID THEN
        alarm_hold := FALSE;
    ELSIF alarm_timer.Q THEN
        alarm_hold := FALSE;
    END_IF;

    alarm_timer(IN := THICKNESS_SIGNAL_VALID AND NOT THICKNESS_FAULT, PT := T#500MS);

    THICKNESS_ALARM := THICKNESS_SIGNAL_VALID AND (valid_fault OR alarm_hold);

    IF THICKNESS_SIGNAL_VALID AND CUTTING_RUN AND NOT THICKNESS_FAULT AND (CycleTime > T#0ms) THEN
        Slab_Runtime_Accumulator := Slab_Runtime_Accumulator + TO_LTIME(CycleTime);
    END_IF;
END_IF;
END_FUNCTION_BLOCK

(* ---- public-medium-06.raw_candidate_02.st ---- *)
(* ENGINEERING_CONTRACT
   THICKNESS_ALARM: latch on valid-fault FALSE->TRUE edge; hold via alarm_hold until TON reaches PT after fault deassert;
   clear on signal invalid; output = signal valid AND alarm_hold; PUB001/PUB004. Current TON.Q read after call.
   Slab_Fault_Counter: increment on same edge; wrap at UINT natural boundary; PUB002/PUB005.
   Slab_Runtime_Accumulator: add TO_LTIME(CycleTime) when valid and CUTTING_RUN and no fault and CycleTime>0 including first scan; LTIME ns; PUB003/PUB004.
   Slab_Fault_History[0..4]: shift oldest right, store timestamp at index0; PUB002/PUB006.
   Power-up: clear all stored state then process current inputs; prev_valid_fault starts false so first valid fault is a transition; PUB005.
   Unspecified: initial fault + invalid signal keeps alarm off until next edge; PUB004/PUB006.
*)
(* CONTRACT_RULES [] *)
FUNCTION_BLOCK SlabThicknessAlarmFaultHistory
VAR_INPUT
    THICKNESS_FAULT : BOOL;
    THICKNESS_SIGNAL_VALID : BOOL;
    CUTTING_RUN : BOOL;
    FaultTimestamp : DINT;
    CycleTime : TIME;
END_VAR
VAR_OUTPUT
    THICKNESS_ALARM : BOOL;
    Slab_Fault_Counter : UINT;
    Slab_Runtime_Accumulator : LTIME;
    Slab_Fault_History : ARRAY[0..4] OF DINT;
END_VAR
VAR
    alarm_hold : BOOL := FALSE;
    alarm_timer : TON;
    prev_valid_fault : BOOL := FALSE;
    init_done : BOOL := FALSE;
    valid_fault : BOOL;
END_VAR

valid_fault := THICKNESS_SIGNAL_VALID AND THICKNESS_FAULT;

IF NOT init_done THEN
    init_done := TRUE;
    Slab_Fault_Counter := UINT#0;
    Slab_Runtime_Accumulator := LTIME#0s;
    Slab_Fault_History[0] := DINT#0;
    Slab_Fault_History[1] := DINT#0;
    Slab_Fault_History[2] := DINT#0;
    Slab_Fault_History[3] := DINT#0;
    Slab_Fault_History[4] := DINT#0;
    alarm_hold := FALSE;
    alarm_timer(IN := FALSE, PT := T#500MS);
    THICKNESS_ALARM := FALSE;
END_IF;

IF valid_fault AND NOT prev_valid_fault THEN
    Slab_Fault_History[4] := Slab_Fault_History[3];
    Slab_Fault_History[3] := Slab_Fault_History[2];
    Slab_Fault_History[2] := Slab_Fault_History[1];
    Slab_Fault_History[1] := Slab_Fault_History[0];
    Slab_Fault_History[0] := FaultTimestamp;
    Slab_Fault_Counter := Slab_Fault_Counter + UINT#1;
    alarm_hold := TRUE;
END_IF;

prev_valid_fault := valid_fault;

alarm_timer(IN := THICKNESS_SIGNAL_VALID AND NOT THICKNESS_FAULT, PT := T#500MS);

IF NOT THICKNESS_SIGNAL_VALID THEN
    alarm_hold := FALSE;
ELSIF NOT valid_fault AND alarm_timer.Q THEN
    alarm_hold := FALSE;
END_IF;

THICKNESS_ALARM := THICKNESS_SIGNAL_VALID AND alarm_hold;

IF THICKNESS_SIGNAL_VALID AND CUTTING_RUN AND NOT THICKNESS_FAULT AND (CycleTime > T#0ms) THEN
    Slab_Runtime_Accumulator := Slab_Runtime_Accumulator + TO_LTIME(CycleTime);
END_IF;

END_FUNCTION_BLOCK

(* ---- public-medium-07.candidate_01.st ---- *)
FUNCTION_BLOCK OfficeHVACMultiModeControl

(* ENGINEERING_CONTRACT
PUB001: HVAC_MODE_SELECTOR valid 0..3; assumption: input is valid.
PUB002: SUPPLY_FAN_RUN active when OCCUPANCY_DETECTED AND mode<>3 remain true for 30s via TON.
  Activation: TON.Q after 30s; Hold: conditions remain true; Reset: occupancy lost or mode=3,
  timer IN false => immediate Q false and ET reset; same-scan final value from current inputs.
PUB003-PUB005: TEMP_SETPOINT_ADJUST combinational from current mode, occupancy, energy-saving.
  Auto: occ 0, unocc ES +3, unocc std +2. Comfort: occ 0, unocc +1.
  Economy: occ 0, unocc +4. Night: +4 regardless of occupancy. Units degrees C.
  Clamp -4..+4. Energy-saving affects Auto mode only.
PUB006: outputs initialized FALSE/0 by declaration/start scan; no independent retained output outside timer.
PUB007: 30s delay controls only BOOL fan enable.
*)

(* CONTRACT_RULES
[]
*)

VAR
    tmp_delayActive : BOOL;
    tmp_fanTimer    : TON;
    tmp_adjust      : INT;
    tmp_mode        : INT;
    tmp_occ         : BOOL;
    tmp_es          : BOOL;
END_VAR

SUPPLY_FAN_RUN := FALSE;
TEMP_SETPOINT_ADJUST := 0;

tmp_mode := HVAC_MODE_SELECTOR;
tmp_occ  := OCCUPANCY_DETECTED;
tmp_es   := ENERGY_SAVING_MODE;

tmp_delayActive := tmp_occ AND (tmp_mode <> 3);
tmp_fanTimer(IN := tmp_delayActive, PT := T#30S);
SUPPLY_FAN_RUN := tmp_fanTimer.Q;

CASE tmp_mode OF
  0:
    IF tmp_occ THEN
      tmp_adjust := 0;
    ELSE
      IF tmp_es THEN
        tmp_adjust := 3;
      ELSE
        tmp_adjust := 2;
      END_IF;
    END_IF;

  1:
    IF tmp_occ THEN
      tmp_adjust := 0;
    ELSE
      tmp_adjust := 1;
    END_IF;

  2:
    IF tmp_occ THEN
      tmp_adjust := 0;
    ELSE
      tmp_adjust := 4;
    END_IF;

  3:
    tmp_adjust := 4;

  ELSE
    tmp_adjust := 0;
END_CASE;

IF tmp_adjust > 4 THEN
  tmp_adjust := 4;
ELSIF tmp_adjust < -4 THEN
  tmp_adjust := -4;
END_IF;

TEMP_SETPOINT_ADJUST := tmp_adjust;

END_FUNCTION_BLOCK

(* ---- public-medium-07.candidate_02.st ---- *)
FUNCTION_BLOCK OfficeHVACMultiModeControl

(* ENGINEERING_CONTRACT
PUB001: HVAC_MODE_SELECTOR valid 0..3; assumption: input is valid.
PUB002: SUPPLY_FAN_RUN active when OCCUPANCY_DETECTED AND mode<>3 remain true for 30s via TON.
  Activation: TON.Q after 30s; Hold: conditions remain true; Reset: occupancy lost or mode=3,
  timer IN false => immediate Q false and ET reset; same-scan final value from current inputs.
PUB003-PUB005: TEMP_SETPOINT_ADJUST combinational from current mode, occupancy, energy-saving.
  Auto: occ 0, unocc ES +3, unocc std +2. Comfort: occ 0, unocc +1.
  Economy: occ 0, unocc +4. Night: +4 regardless of occupancy. Units degrees C.
  Clamp -4..+4. Energy-saving affects Auto mode only.
PUB006: outputs initialized FALSE/0 by declaration/start scan; no independent retained output outside timer.
PUB007: 30s delay controls only BOOL fan enable.
*)

(* CONTRACT_RULES
[]
*)

VAR_INPUT
    OCCUPANCY_DETECTED : BOOL;
    ENERGY_SAVING_MODE : BOOL;
    HVAC_MODE_SELECTOR : INT;
END_VAR
VAR_OUTPUT
    SUPPLY_FAN_RUN : BOOL;
    TEMP_SETPOINT_ADJUST : INT;
END_VAR
VAR
    tmp_delayActive : BOOL;
    tmp_fanTimer    : TON;
    tmp_adjust      : INT;
    tmp_mode        : INT;
    tmp_occ         : BOOL;
    tmp_es          : BOOL;
END_VAR

SUPPLY_FAN_RUN := FALSE;
TEMP_SETPOINT_ADJUST := 0;

tmp_mode := HVAC_MODE_SELECTOR;
tmp_occ  := OCCUPANCY_DETECTED;
tmp_es   := ENERGY_SAVING_MODE;

tmp_delayActive := tmp_occ AND (tmp_mode <> 3);
tmp_fanTimer(IN := tmp_delayActive, PT := T#30S);
SUPPLY_FAN_RUN := tmp_fanTimer.Q;

CASE tmp_mode OF
  0:
    IF tmp_occ THEN
      tmp_adjust := 0;
    ELSE
      IF tmp_es THEN
        tmp_adjust := 3;
      ELSE
        tmp_adjust := 2;
      END_IF;
    END_IF;

  1:
    IF tmp_occ THEN
      tmp_adjust := 0;
    ELSE
      tmp_adjust := 1;
    END_IF;

  2:
    IF tmp_occ THEN
      tmp_adjust := 0;
    ELSE
      tmp_adjust := 4;
    END_IF;

  3:
    tmp_adjust := 4;

  ELSE
    tmp_adjust := 0;
END_CASE;

IF tmp_adjust > 4 THEN
  tmp_adjust := 4;
ELSIF tmp_adjust < -4 THEN
  tmp_adjust := -4;
END_IF;

TEMP_SETPOINT_ADJUST := tmp_adjust;

END_FUNCTION_BLOCK

(* ---- public-medium-07.raw_candidate_01.st ---- *)
FUNCTION_BLOCK OfficeHVACMultiModeControl

(* ENGINEERING_CONTRACT
PUB001: HVAC_MODE_SELECTOR valid 0..3; assumption: input is valid.
PUB002: SUPPLY_FAN_RUN active when OCCUPANCY_DETECTED AND mode<>3 remain true for 30s via TON.
  Activation: TON.Q after 30s; Hold: conditions remain true; Reset: occupancy lost or mode=3,
  timer IN false => immediate Q false and ET reset; same-scan final value from current inputs.
PUB003-PUB005: TEMP_SETPOINT_ADJUST combinational from current mode, occupancy, energy-saving.
  Auto: occ 0, unocc ES +3, unocc std +2. Comfort: occ 0, unocc +1.
  Economy: occ 0, unocc +4. Night: +4 regardless of occupancy. Units degrees C.
  Clamp -4..+4. Energy-saving affects Auto mode only.
PUB006: outputs initialized FALSE/0 by declaration/start scan; no independent retained output outside timer.
PUB007: 30s delay controls only BOOL fan enable.
*)

(* CONTRACT_RULES
[]
*)

VAR
    tmp_delayActive : BOOL;
    tmp_fanTimer    : TON;
    tmp_adjust      : INT;
    tmp_mode        : INT;
    tmp_occ         : BOOL;
    tmp_es          : BOOL;
END_VAR

SUPPLY_FAN_RUN := FALSE;
TEMP_SETPOINT_ADJUST := 0;

tmp_mode := HVAC_MODE_SELECTOR;
tmp_occ  := OCCUPANCY_DETECTED;
tmp_es   := ENERGY_SAVING_MODE;

tmp_delayActive := tmp_occ AND (tmp_mode <> 3);
tmp_fanTimer(IN := tmp_delayActive, PT := T#30S);
SUPPLY_FAN_RUN := tmp_fanTimer.Q;

CASE tmp_mode OF
  0:
    IF tmp_occ THEN
      tmp_adjust := 0;
    ELSE
      IF tmp_es THEN
        tmp_adjust := 3;
      ELSE
        tmp_adjust := 2;
      END_IF;
    END_IF;

  1:
    IF tmp_occ THEN
      tmp_adjust := 0;
    ELSE
      tmp_adjust := 1;
    END_IF;

  2:
    IF tmp_occ THEN
      tmp_adjust := 0;
    ELSE
      tmp_adjust := 4;
    END_IF;

  3:
    tmp_adjust := 4;

  ELSE
    tmp_adjust := 0;
END_CASE;

IF tmp_adjust > 4 THEN
  tmp_adjust := 4;
ELSIF tmp_adjust < -4 THEN
  tmp_adjust := -4;
END_IF;

TEMP_SETPOINT_ADJUST := tmp_adjust;

END_FUNCTION_BLOCK

(* ---- public-medium-07.raw_candidate_02.st ---- *)
FUNCTION_BLOCK OfficeHVACMultiModeControl

(* ENGINEERING_CONTRACT
PUB001: HVAC_MODE_SELECTOR valid 0..3; assumption: input is valid.
PUB002: SUPPLY_FAN_RUN active when OCCUPANCY_DETECTED AND mode<>3 remain true for 30s via TON.
  Activation: TON.Q after 30s; Hold: conditions remain true; Reset: occupancy lost or mode=3,
  timer IN false => immediate Q false and ET reset; same-scan final value from current inputs.
PUB003-PUB005: TEMP_SETPOINT_ADJUST combinational from current mode, occupancy, energy-saving.
  Auto: occ 0, unocc ES +3, unocc std +2. Comfort: occ 0, unocc +1.
  Economy: occ 0, unocc +4. Night: +4 regardless of occupancy. Units degrees C.
  Clamp -4..+4. Energy-saving affects Auto mode only.
PUB006: outputs initialized FALSE/0 by declaration/start scan; no independent retained output outside timer.
PUB007: 30s delay controls only BOOL fan enable.
*)

(* CONTRACT_RULES
[]
*)

VAR_INPUT
    OCCUPANCY_DETECTED : BOOL;
    ENERGY_SAVING_MODE : BOOL;
    HVAC_MODE_SELECTOR : INT;
END_VAR
VAR_OUTPUT
    SUPPLY_FAN_RUN : BOOL;
    TEMP_SETPOINT_ADJUST : INT;
END_VAR
VAR
    tmp_delayActive : BOOL;
    tmp_fanTimer    : TON;
    tmp_adjust      : INT;
    tmp_mode        : INT;
    tmp_occ         : BOOL;
    tmp_es          : BOOL;
END_VAR

SUPPLY_FAN_RUN := FALSE;
TEMP_SETPOINT_ADJUST := 0;

tmp_mode := HVAC_MODE_SELECTOR;
tmp_occ  := OCCUPANCY_DETECTED;
tmp_es   := ENERGY_SAVING_MODE;

tmp_delayActive := tmp_occ AND (tmp_mode <> 3);
tmp_fanTimer(IN := tmp_delayActive, PT := T#30S);
SUPPLY_FAN_RUN := tmp_fanTimer.Q;

CASE tmp_mode OF
  0:
    IF tmp_occ THEN
      tmp_adjust := 0;
    ELSE
      IF tmp_es THEN
        tmp_adjust := 3;
      ELSE
        tmp_adjust := 2;
      END_IF;
    END_IF;

  1:
    IF tmp_occ THEN
      tmp_adjust := 0;
    ELSE
      tmp_adjust := 1;
    END_IF;

  2:
    IF tmp_occ THEN
      tmp_adjust := 0;
    ELSE
      tmp_adjust := 4;
    END_IF;

  3:
    tmp_adjust := 4;

  ELSE
    tmp_adjust := 0;
END_CASE;

IF tmp_adjust > 4 THEN
  tmp_adjust := 4;
ELSIF tmp_adjust < -4 THEN
  tmp_adjust := -4;
END_IF;

TEMP_SETPOINT_ADJUST := tmp_adjust;

END_FUNCTION_BLOCK

(* ---- public-medium-08.candidate_01.st ---- *)
(* ENGINEERING_CONTRACT
   ipValue: combinational output from current ipText; no retained/latched state.
   Activation: exactly 4 non-empty decimal segments, each value 0..255
   (PUB001, PUB003). Assemble network byte order (PUB002).
   Zero/deactivation: malformed, non-digit, wrong segment count, out-of-range,
   empty/short (<7), or length >15 characters (PUB003, PUB004).
   0.0.0.0 also produces 0.
   Same-scan: input is read once per call; no priority or reset inputs.
   Boundaries: first segment bits31..24, second bits23..16, third bits15..8,
   fourth bits7..0; UDINT result.
 *)
(* CONTRACT_RULES [] *)
FUNCTION_BLOCK IPv4Parser
VAR_INPUT
    ipText : STRING(254);
END_VAR
VAR_OUTPUT
    ipValue : UDINT;
END_VAR
VAR
    tmp_len : INT;
    tmp_i : INT;
    tmp_ch : BYTE;
    tmp_segVal : UDINT;
    tmp_segCount : INT;
    tmp_digitCount : INT;
    tmp_addr : UDINT;
END_VAR

ipValue := UDINT#0;

tmp_len := LEN(ipText);
IF (tmp_len < 7) OR (tmp_len > 15) THEN
    RETURN;
END_IF;

tmp_segVal := UDINT#0;
tmp_segCount := 0;
tmp_digitCount := 0;
tmp_addr := UDINT#0;

FOR tmp_i := 0 TO (tmp_len - 1) DO
    tmp_ch := ipText[tmp_i];

    IF (tmp_ch >= BYTE#48) AND (tmp_ch <= BYTE#57) THEN
        tmp_digitCount := tmp_digitCount + 1;
        tmp_segVal := (tmp_segVal * UDINT#10) + (BYTE_TO_UDINT(tmp_ch) - UDINT#48);
        IF tmp_segVal > UDINT#255 THEN
            RETURN;
        END_IF;
    ELSIF tmp_ch = BYTE#46 THEN
        IF tmp_digitCount = 0 THEN
            RETURN;
        END_IF;
        IF tmp_segCount >= 3 THEN
            RETURN;
        END_IF;

        tmp_addr := SHL(tmp_addr, 8);
        tmp_addr := tmp_addr OR (tmp_segVal AND UDINT#255);

        tmp_segCount := tmp_segCount + 1;
        tmp_segVal := UDINT#0;
        tmp_digitCount := 0;
    ELSE
        RETURN;
    END_IF;
END_FOR;

IF (tmp_digitCount = 0) OR (tmp_segCount <> 3) THEN
    RETURN;
END_IF;

tmp_addr := SHL(tmp_addr, 8);
tmp_addr := tmp_addr OR (tmp_segVal AND UDINT#255);
ipValue := tmp_addr;

END_FUNCTION_BLOCK

(* ---- public-medium-08.raw_candidate_01.st ---- *)
(* ENGINEERING_CONTRACT
   ipValue: combinational output from current ipText; no retained/latched state.
   Activation: exactly 4 non-empty decimal segments, each value 0..255
   (PUB001, PUB003). Assemble network byte order (PUB002).
   Zero/deactivation: malformed, non-digit, wrong segment count, out-of-range,
   empty/short (<7), or length >15 characters (PUB003, PUB004).
   0.0.0.0 also produces 0.
   Same-scan: input is read once per call; no priority or reset inputs.
   Boundaries: first segment bits31..24, second bits23..16, third bits15..8,
   fourth bits7..0; UDINT result.
 *)
(* CONTRACT_RULES [] *)
FUNCTION_BLOCK IPv4Parser
VAR_INPUT
    ipText : STRING(254);
END_VAR
VAR_OUTPUT
    ipValue : UDINT;
END_VAR
VAR
    tmp_len : INT;
    tmp_i : INT;
    tmp_ch : BYTE;
    tmp_segVal : UDINT;
    tmp_segCount : INT;
    tmp_digitCount : INT;
    tmp_addr : UDINT;
END_VAR

ipValue := UDINT#0;

tmp_len := LEN(ipText);
IF (tmp_len < 7) OR (tmp_len > 15) THEN
    RETURN;
END_IF;

tmp_segVal := UDINT#0;
tmp_segCount := 0;
tmp_digitCount := 0;
tmp_addr := UDINT#0;

FOR tmp_i := 0 TO (tmp_len - 1) DO
    tmp_ch := ipText[tmp_i];

    IF (tmp_ch >= BYTE#48) AND (tmp_ch <= BYTE#57) THEN
        tmp_digitCount := tmp_digitCount + 1;
        tmp_segVal := (tmp_segVal * UDINT#10) + (BYTE_TO_UDINT(tmp_ch) - UDINT#48);
        IF tmp_segVal > UDINT#255 THEN
            RETURN;
        END_IF;
    ELSIF tmp_ch = BYTE#46 THEN
        IF tmp_digitCount = 0 THEN
            RETURN;
        END_IF;
        IF tmp_segCount >= 3 THEN
            RETURN;
        END_IF;

        tmp_addr := SHL(tmp_addr, 8);
        tmp_addr := tmp_addr OR (tmp_segVal AND UDINT#255);

        tmp_segCount := tmp_segCount + 1;
        tmp_segVal := UDINT#0;
        tmp_digitCount := 0;
    ELSE
        RETURN;
    END_IF;
END_FOR;

IF (tmp_digitCount = 0) OR (tmp_segCount <> 3) THEN
    RETURN;
END_IF;

tmp_addr := SHL(tmp_addr, 8);
tmp_addr := tmp_addr OR (tmp_segVal AND UDINT#255);
ipValue := tmp_addr;

END_FUNCTION_BLOCK
